DATA_BLOCK "db3202_BC595_SetupPorTensao"
TITLE = db3202_BC595_SetupPorTensao v0.2 (DB3202)
{ S7_Optimized_Access := 'FALSE' }
AUTHOR : 'Reginaldo Lobo'
VERSION : 0.2
////====================================
//// db3202_BC595_SetupPorTensao (DB3202) - GERADO por plc/bt2/gerador/gerar_banco_v0.2.py (03/11/2026) - nao compilado, nao testado
//// O QUE FAZ : mesmo papel do db152_BC56_SetupPorTensao v0.2, 32 chaves por chaveamento (1=220, 2=380, 3=440 V). Banco BC59,5.
//// p = (chaveamento-1)*32 + (chave-1)  (0..95)
//// OFFSETS (calculados; CONFERIR no TIA): tensaoV W0/2/4 | kwReal D6+4p | rMedidoOhm D390+4p | vMedidaV D774+4p
////    baseKw D1158+4p | setupData B1542+12p | setupOk X2694.0+p | selV.tensaoSel W2706
//// RETENTIVIDADE : precisa sobreviver a reinicio da CPU; conferir no TIA.
////=====================================
   VAR
      setupV : Struct
         tensaoV     : Array[1..3] of Int;
         kwReal      : Array[1..3, 1..32] of Real;
         rMedidoOhm  : Array[1..3, 1..32] of Real;
         vMedidaV    : Array[1..3, 1..32] of Real;
         baseKw      : Array[1..3, 1..32] of Real;
         setupData   : Array[1..3, 1..32] of DTL;
         setupOk     : Array[1..3, 1..32] of Bool;
      END_STRUCT;
      selV : Struct
         tensaoSel   : Int;
      END_STRUCT;
   END_VAR


BEGIN
   setupV.tensaoV[1] := 220;
   setupV.tensaoV[2] := 380;
   setupV.tensaoV[3] := 440;
   selV.tensaoSel := 0;   // NAO informado ate o operador escolher no HTML

END_DATA_BLOCK
